(* IEC 61131-3 sources: Versio-VersionControlSystem/fixtures/projects/TC3_PlcSample_reStrText/TC3_PlcSample_reStrText/LibraryDocumentationSample Project/LibPOUs/B_DocuElements/Internal Comments, 1 file *)

(* ---- FB_Libdoc_InternalComments.st ---- *)
(*
This is the first paragraph.

.. Comments begin with two dots and one space. Anything can
   follow, except for the syntax of footnotes/citations,
   hyperlink targets, directives, or substitution definitions.

Since comments are not shown, this paragraph follows the previous paragraph directly.
*)

FUNCTION_BLOCK FB_Libdoc_InternalComments
VAR_INPUT
    nVarA : INT;
    nVarB : INT;
END_VAR
VAR_OUTPUT
    nSum : INT;
END_VAR
VAR
END_VAR
